Fanuc KAREL source: KB00094.KL

PROGRAM KB00094
%NOLOCKGROUP
%ENVIRONMENT TIM
VAR
  P1: INTEGER
BEGIN
  P1 = 1
  GET_TIME(P1)
END KB00094
